(* IEC 61131-3 sources: SortJet_MasterSPS_Aufbau.fbsproj/Device.device.xml.v3^/Plc Logic.plclogic.xml.v3^/Application.application.xml.v3^/09_Station/Shuttle/[101,102] Shuttle/0_Konfig (part 2) *)

(* ---- Konfiguration_101.gvl ---- *)
(* METADATA
{
	"v3Meta": {
		"objectGuid": "a708fc7a-282c-4202-ac62-7eb4c755f260"
	}
}
*)
{attribute 'allow_unqualified_access'}
NAMESPACE Konfiguration_101
VAR_CONFIG
  // werden Variablen die gemappt werden hier ignoriert?
  // ------------------------------------------------- HARDWARE EINGAENGE -------------------------------------------------
  // Datenlichtschranke
  Globale_Bausteine.aShuttle[101].in_bDatenlichtschrankeShuttlebahnOK                                AT %MX1.1  : BOOL; // OPTION - Bauteil an der Shuttlebahn => Sender / Empfaenger
  Globale_Bausteine.aShuttle[101].in_bDatenlichtschrankeShuttleOK                                    AT %MX1.1  : BOOL; // OPTION - Bauteil auf dem Shuttle => Sender / Empfaenger

  // Sicherungen \ Motorschutzschalter \ etc.

  Globale_Bausteine.aShuttle[101].in_bSicherungen230V_OK                                             AT %MX1.1   : BOOL; // OPTION
  Globale_Bausteine.aShuttle[101].in_bLSQuerfahrtBremseOK                                            AT %IX101.0 : BOOL; // IO-L - Querfahrt Bremse Sicherung
  Globale_Bausteine.aShuttle[101].in_bNetzteil_24V_OK                                                AT %IX100.1 : BOOL; // IO-L - Netzteil 24V OK
  Globale_Bausteine.aShuttle[101].Kippen.in_bLeitungsschutzschalterBremseOK                          AT %MX1.1   : BOOL; // OPTION
  Globale_Bausteine.aShuttle[101].Kippen.in_bMotorschutzschalter_OK                                  AT %MX1.1   : BOOL; // OPTION

  // Druckluft
  Globale_Bausteine.aShuttle[101].in_bSicherungKompressor_OK                                         AT %MX1.1  : BOOL; // OPTION
  Globale_Bausteine.aShuttle[101].in_bDruckluft_OK                                                   AT %MX1.1  : BOOL; // OPTION

  //Geblaese Wand 1
  Globale_Bausteine.aShuttle[101].Geblaese[1].in_bMotorschutzschalter_OK                             AT %IX101.1  : BOOL; // IO-L - Geblaesegruppe Wand 1 Sicherung + Motorschutz
  Globale_Bausteine.aShuttle[101].Geblaese[1].out_bStarteGeblaese                                    AT %QX100.1  : BOOL; // IO-L - Geblaesegruppe Wand 1 einschalten

  // Wandverstellung Wand 1
  Globale_Bausteine.aShuttle[101].in_bWandverstellungsAntriebsSicherungOK                            AT %MX1.1   : BOOL; // OPTION
  Globale_Bausteine.aShuttle[101].in_bMotorstarterWandverstellungOK                                  AT %MX1.1   : BOOL; // OPTION
  Globale_Bausteine.aShuttle[101].in_bWandverstellungsBremsSicherungOK                               AT %MX1.1   : BOOL; // OPTION

  Globale_Bausteine.aShuttle[101].Wandverstellung[1].Pneumatik.in_bWandEinlaufseiteGeoeffnet         AT %MX1.0   : BOOL; // OPTION
  Globale_Bausteine.aShuttle[101].Wandverstellung[1].Pneumatik.in_bWandEinlaufseiteGeschlossen       AT %MX1.0   : BOOL; // OPTION
  Globale_Bausteine.aShuttle[101].Wandverstellung[1].Pneumatik.in_bWandAuslaufseiteGeoeffnet         AT %MX1.0   : BOOL; // OPTION
  Globale_Bausteine.aShuttle[101].Wandverstellung[1].Pneumatik.in_bWandAuslaufseiteGeschlossen       AT %MX1.0   : BOOL; // OPTION

  Globale_Bausteine.aShuttle[101].Wandverstellung[1].Pneumatik.out_bWandverstellungOeffnen           AT %MX1010.1 : BOOL; // OPTION
  Globale_Bausteine.aShuttle[101].Wandverstellung[1].Pneumatik.out_bWandverstellungSchliessen        AT %MX1010.2 : BOOL; // OPTION

  Globale_Bausteine.aShuttle[101].Wandverstellung[1].Pneumatik2.in_bStatusZylinder_Alle_Eingefahren  AT %MX1.0   : BOOL; // OPTION
  Globale_Bausteine.aShuttle[101].Wandverstellung[1].Pneumatik2.in_bStatusZylinder_1_Ausgefahren     AT %MX1.0   : BOOL; // OPTION
  Globale_Bausteine.aShuttle[101].Wandverstellung[1].Pneumatik2.in_bStatusZylinder_2_Ausgefahren     AT %MX1.0   : BOOL; // OPTION

  Globale_Bausteine.aShuttle[101].Wandverstellung[1].Pneumatik2.out_bZylinder_1_Einfahren            AT %MX1010.3 : BOOL; // OPTION
  Globale_Bausteine.aShuttle[101].Wandverstellung[1].Pneumatik2.out_bZylinder_2_Einfahren            AT %MX1010.4 : BOOL; // OPTION
  Globale_Bausteine.aShuttle[101].Wandverstellung[1].Pneumatik2.out_bZylinder_1_Ausfahren            AT %MX1010.5 : BOOL; // OPTION
  Globale_Bausteine.aShuttle[101].Wandverstellung[1].Pneumatik2.out_bZylinder_2_Ausfahren            AT %MX1010.6 : BOOL; // OPTION

  Globale_Bausteine.aShuttle[101].Wandverstellung[1].Rollenleiste.in_bStatusZylinder1Ausgefahren     AT %MX1.0   : BOOL; // OPTION
  Globale_Bausteine.aShuttle[101].Wandverstellung[1].Rollenleiste.in_bStatusZylinder1Eingefahren     AT %MX1.0   : BOOL; // OPTION
  Globale_Bausteine.aShuttle[101].Wandverstellung[1].Rollenleiste.in_bStatusZylinder2Ausgefahren     AT %MX1.0   : BOOL; // OPTION
  Globale_Bausteine.aShuttle[101].Wandverstellung[1].Rollenleiste.in_bStatusZylinder2Eingefahren     AT %MX1.0   : BOOL; // OPTION

  Globale_Bausteine.aShuttle[101].Wandverstellung[1].Rollenleiste.out_bZylinder1Einfahren            AT %MX1010.7 : BOOL; // OPTION
  Globale_Bausteine.aShuttle[101].Wandverstellung[1].Rollenleiste.out_bZylinder1Ausfahren            AT %MX1011.0 : BOOL; // OPTION
  Globale_Bausteine.aShuttle[101].Wandverstellung[1].Rollenleiste.out_bZylinder2Einfahren            AT %MX1011.1 : BOOL; // OPTION
  Globale_Bausteine.aShuttle[101].Wandverstellung[1].Rollenleiste.out_bZylinder2Ausfahren            AT %MX1011.2 : BOOL; // OPTION

  Globale_Bausteine.aShuttle[101].Wandverstellung[1].Rollenleiste_Schuetz.in_bVerstellungGeoeffnet   AT %MX1.0   : BOOL; // OPTION
  Globale_Bausteine.aShuttle[101].Wandverstellung[1].Rollenleiste_Schuetz.in_bVerstellungGeschlossen AT %MX1.0   : BOOL; // OPTION
  Globale_Bausteine.aShuttle[101].Wandverstellung[1].Rollenleiste_Schuetz.in_bMotorstarter_OK        AT %MX1.1   : BOOL; // OPTION
  Globale_Bausteine.aShuttle[101].Wandverstellung[1].Rollenleiste_Schuetz.in_bSicherungMotorOK       AT %MX1.1   : BOOL; // OPTION
  Globale_Bausteine.aShuttle[101].Wandverstellung[1].Rollenleiste_Schuetz.in_bBremseOK               AT %MX1.1   : BOOL; // OPTION

  Globale_Bausteine.aShuttle[101].Wandverstellung[1].Rollenleiste_Schuetz.out_bVerstellungSchliessen AT %MX1011.3 : BOOL; // OPTION
  Globale_Bausteine.aShuttle[101].Wandverstellung[1].Rollenleiste_Schuetz.out_bVerstellungOeffnen    AT %MX1011.4 : BOOL; // OPTION
  Globale_Bausteine.aShuttle[101].Wandverstellung[1].Rollenleiste_Schuetz.out_bBremseOeffnen         AT %MX1011.5 : BOOL; // OPTION
  Globale_Bausteine.aShuttle[101].Wandverstellung[1].Rollenleiste_Schuetz.out_bMotorstarterReset     AT %MX1011.6 : BOOL; // OPTION

  Globale_Bausteine.aShuttle[101].Wandverstellung[1].Gegenhalter_Schuetz.in_bVerstellungGeoeffnet    AT %MX1.0   : BOOL; // OPTION
  Globale_Bausteine.aShuttle[101].Wandverstellung[1].Gegenhalter_Schuetz.in_bVerstellungGeschlossen  AT %MX1.0   : BOOL; // OPTION
  Globale_Bausteine.aShuttle[101].Wandverstellung[1].Gegenhalter_Schuetz.in_bMotorstarter_OK         AT %MX1.1   : BOOL; // OPTION
  Globale_Bausteine.aShuttle[101].Wandverstellung[1].Gegenhalter_Schuetz.in_bSicherungMotorOK        AT %MX1.1   : BOOL; // OPTION
  Globale_Bausteine.aShuttle[101].Wandverstellung[1].Gegenhalter_Schuetz.in_bBremseOK                AT %MX1.1   : BOOL; // OPTION

  Globale_Bausteine.aShuttle[101].Wandverstellung[1].Gegenhalter_Schuetz.out_bVerstellungSchliessen  AT %MX1011.7 : BOOL; // OPTION
  Globale_Bausteine.aShuttle[101].Wandverstellung[1].Gegenhalter_Schuetz.out_bVerstellungOeffnen     AT %MX1012.0 : BOOL; // OPTION
  Globale_Bausteine.aShuttle[101].Wandverstellung[1].Gegenhalter_Schuetz.out_bBremseOeffnen          AT %MX1012.1 : BOOL; // OPTION
  Globale_Bausteine.aShuttle[101].Wandverstellung[1].Gegenhalter_Schuetz.out_bMotorstarterReset      AT %MX1012.2 : BOOL; // OPTION

  // Sensoren  Wand 2
  Globale_Bausteine.aShuttle[101].in_bSensorEinlaufVorabWand2                                        AT %MX1.0   : BOOL; // OPTION
  Globale_Bausteine.aShuttle[101].in_bSensorAuslaufVorabWand2                                        AT %MX1.0   : BOOL; // OPTION
  Globale_Bausteine.aShuttle[101].in_bSensorAuslaufStoppWand2                                        AT %MX1.0   : BOOL; // OPTION

  // Greifer Wand 1 [Ausbaustufe stStationsAufbau.bGreifer] (Kanaele laut Schaltplan eintragen, Glasrueckhalter laut Parameter_Greifer, ohne Bauteil Eingang auf %MX1.1)
  Globale_Bausteine.aShuttle[101].Greifer[1].in_bGreiferAusgefahren                                     AT %MX1.0   : BOOL; // OPTION
  Globale_Bausteine.aShuttle[101].Greifer[1].in_bGreiferEingefahren                                     AT %MX1.0   : BOOL; // OPTION
  Globale_Bausteine.aShuttle[101].Greifer[1].in_bGlasRueckhalterEinlaufEingefahren                      AT %MX1.1   : BOOL; // OPTION
  Globale_Bausteine.aShuttle[101].Greifer[1].in_bGlasRueckhalterAuslaufEingefahren                      AT %MX1.1   : BOOL; // OPTION

  Globale_Bausteine.aShuttle[101].Greifer[1].out_bGreiferAusfahren                                      AT %MX1012.3 : BOOL; // OPTION
  Globale_Bausteine.aShuttle[101].Greifer[1].out_bGreiferEinfahren                                      AT %MX1012.4 : BOOL; // OPTION
  Globale_Bausteine.aShuttle[101].Greifer[1].out_bGlasRueckhalterEinlaufAusfahren                       AT %MX1012.5 : BOOL; // OPTION
  Globale_Bausteine.aShuttle[101].Greifer[1].out_bGlasRueckhalterAuslaufAusfahren                       AT %MX1012.6 : BOOL; // OPTION

  // Greiferzange Einlaufseite Wand 1 [nur mit Parameter_Greifer.bZangeEinlaufVorhanden]
  Globale_Bausteine.aShuttle[101].Greifer[1].Zange[1].in_bStatusZylinder_Alle_Eingefahren               AT %MX1.0   : BOOL; // OPTION
  Globale_Bausteine.aShuttle[101].Greifer[1].Zange[1].in_bStatusZylinder_1_Ausgefahren                  AT %MX1.0   : BOOL; // OPTION
  Globale_Bausteine.aShuttle[101].Greifer[1].Zange[1].in_bStatusZylinder_2_Ausgefahren                  AT %MX1.0   : BOOL; // OPTION
  Globale_Bausteine.aShuttle[101].Greifer[1].Zange[1].in_bStatusZylinder_3_Ausgefahren                  AT %MX1.0   : BOOL; // OPTION

  Globale_Bausteine.aShuttle[101].Greifer[1].Zange[1].out_bZylinder_1_Einfahren                         AT %MX1012.7 : BOOL; // OPTION
  Globale_Bausteine.aShuttle[101].Greifer[1].Zange[1].out_bZylinder_2_Einfahren                         AT %MX1013.0 : BOOL; // OPTION
  Globale_Bausteine.aShuttle[101].Greifer[1].Zange[1].out_bZylinder_3_Einfahren                         AT %MX1013.1 : BOOL; // OPTION
  Globale_Bausteine.aShuttle[101].Greifer[1].Zange[1].out_bZylinder_1_Ausfahren                         AT %MX1013.2 : BOOL; // OPTION
  Globale_Bausteine.aShuttle[101].Greifer[1].Zange[1].out_bZylinder_2_Ausfahren                         AT %MX1013.3 : BOOL; // OPTION
  Globale_Bausteine.aShuttle[101].Greifer[1].Zange[1].out_bZylinder_3_Ausfahren                         AT %MX1013.4 : BOOL; // OPTION

  // Greiferzange Auslaufseite Wand 1 [nur mit Parameter_Greifer.bZangeAuslaufVorhanden]
  Globale_Bausteine.aShuttle[101].Greifer[1].Zange[2].in_bStatusZylinder_Alle_Eingefahren               AT %MX1.0   : BOOL; // OPTION
  Globale_Bausteine.aShuttle[101].Greifer[1].Zange[2].in_bStatusZylinder_1_Ausgefahren                  AT %MX1.0   : BOOL; // OPTION
  Globale_Bausteine.aShuttle[101].Greifer[1].Zange[2].in_bStatusZylinder_2_Ausgefahren                  AT %MX1.0   : BOOL; // OPTION
  Globale_Bausteine.aShuttle[101].Greifer[1].Zange[2].in_bStatusZylinder_3_Ausgefahren                  AT %MX1.0   : BOOL; // OPTION

  Globale_Bausteine.aShuttle[101].Greifer[1].Zange[2].out_bZylinder_1_Einfahren                         AT %MX1013.5 : BOOL; // OPTION
  Globale_Bausteine.aShuttle[101].Greifer[1].Zange[2].out_bZylinder_2_Einfahren                         AT %MX1013.6 : BOOL; // OPTION
  Globale_Bausteine.aShuttle[101].Greifer[1].Zange[2].out_bZylinder_3_Einfahren                         AT %MX1013.7 : BOOL; // OPTION
  Globale_Bausteine.aShuttle[101].Greifer[1].Zange[2].out_bZylinder_1_Ausfahren                         AT %MX1014.0 : BOOL; // OPTION
  Globale_Bausteine.aShuttle[101].Greifer[1].Zange[2].out_bZylinder_2_Ausfahren                         AT %MX1014.1 : BOOL; // OPTION
  Globale_Bausteine.aShuttle[101].Greifer[1].Zange[2].out_bZylinder_3_Ausfahren                         AT %MX1014.2 : BOOL; // OPTION

END_VAR

END_NAMESPACE

(* ---- Konfiguration_102.gvl ---- *)
(* METADATA
{
	"v3Meta": {
		"objectGuid": "12c6a77b-9420-47d5-ba1c-b94e93a145ed"
	}
}
*)
{attribute 'allow_unqualified_access'}
NAMESPACE Konfiguration_102
VAR_CONFIG
  // werden Variablen die gemappt werden hier ignoriert?
  // ------------------------------------------------- HARDWARE EINGAENGE -------------------------------------------------
  // Datenlichtschranke
  Globale_Bausteine.aShuttle[102].in_bDatenlichtschrankeShuttlebahnOK                                AT %MX1.1  : BOOL; // OPTION - Bauteil an der Shuttlebahn => Sender / Empfaenger
  Globale_Bausteine.aShuttle[102].in_bDatenlichtschrankeShuttleOK                                    AT %MX1.1  : BOOL; // OPTION - Bauteil auf dem Shuttle => Sender / Empfaenger

  // Sicherungen \ Motorschutzschalter \ etc.
  Globale_Bausteine.aShuttle[102].in_bSicherungen230V_OK                                             AT %MX1.1    : BOOL; // OPTION
  Globale_Bausteine.aShuttle[102].in_bLSQuerfahrtBremseOK                                            AT %IX111.0  : BOOL; // IO-L - Querfahrt Bremse Sicherung
  Globale_Bausteine.aShuttle[102].in_bNetzteil_24V_OK                                                AT %IX110.1  : BOOL; // IO-L - Netzteil 24V OK

  Globale_Bausteine.aShuttle[102].Kippen.in_bMotorschutzschalter_OK                                  AT %MX1.1   : BOOL; // OPTION
  Globale_Bausteine.aShuttle[102].Kippen.in_bLeitungsschutzschalterBremseOK                          AT %MX1.1   : BOOL; // OPTION

  // Druckluft
  Globale_Bausteine.aShuttle[102].in_bSicherungKompressor_OK                                         AT %MX1.1   : BOOL; // OPTION
  Globale_Bausteine.aShuttle[102].in_bDruckluft_OK                                                   AT %IX114.5 : BOOL; // IO-L - Druckluft OK

  //Geblaese Wand 1
  Globale_Bausteine.aShuttle[102].Geblaese[1].in_bMotorschutzschalter_OK                             AT %IX111.1  : BOOL; // IO-L - Geblaesegruppe Wand 1 Sicherung + Motorschutz
  Globale_Bausteine.aShuttle[102].Geblaese[1].out_bStarteGeblaese                                    AT %QX110.1  : BOOL; // IO-L - Geblaesegruppe Wand 1 einschalten

  // Wandverstellung Wand 1
  Globale_Bausteine.aShuttle[102].in_bWandverstellungsAntriebsSicherungOK                            AT %MX1.1   : BOOL; // OPTION
  Globale_Bausteine.aShuttle[102].in_bMotorstarterWandverstellungOK                                  AT %MX1.1   : BOOL; // OPTION
  Globale_Bausteine.aShuttle[102].in_bWandverstellungsBremsSicherungOK                               AT %MX1.1   : BOOL; // OPTION

  Globale_Bausteine.aShuttle[102].Wandverstellung[1].Pneumatik.in_bWandEinlaufseiteGeoeffnet         AT %MX1.0   : BOOL; // OPTION
  Globale_Bausteine.aShuttle[102].Wandverstellung[1].Pneumatik.in_bWandEinlaufseiteGeschlossen       AT %MX1.0   : BOOL; // OPTION
  Globale_Bausteine.aShuttle[102].Wandverstellung[1].Pneumatik.in_bWandAuslaufseiteGeoeffnet         AT %MX1.0   : BOOL; // OPTION
  Globale_Bausteine.aShuttle[102].Wandverstellung[1].Pneumatik.in_bWandAuslaufseiteGeschlossen       AT %MX1.0   : BOOL; // OPTION

  Globale_Bausteine.aShuttle[102].Wandverstellung[1].Pneumatik.out_bWandverstellungOeffnen           AT %MX1020.1 : BOOL; // OPTION
  Globale_Bausteine.aShuttle[102].Wandverstellung[1].Pneumatik.out_bWandverstellungSchliessen        AT %MX1020.2 : BOOL; // OPTION

  Globale_Bausteine.aShuttle[102].Wandverstellung[1].Pneumatik2.in_bStatusZylinder_Alle_Eingefahren  AT %MX1.0   : BOOL; // OPTION
  Globale_Bausteine.aShuttle[102].Wandverstellung[1].Pneumatik2.in_bStatusZylinder_1_Ausgefahren     AT %MX1.0   : BOOL; // OPTION
  Globale_Bausteine.aShuttle[102].Wandverstellung[1].Pneumatik2.in_bStatusZylinder_2_Ausgefahren     AT %MX1.0   : BOOL; // OPTION

  Globale_Bausteine.aShuttle[102].Wandverstellung[1].Pneumatik2.out_bZylinder_1_Einfahren            AT %MX1020.3 : BOOL; // OPTION
  Globale_Bausteine.aShuttle[102].Wandverstellung[1].Pneumatik2.out_bZylinder_2_Einfahren            AT %MX1020.4 : BOOL; // OPTION
  Globale_Bausteine.aShuttle[102].Wandverstellung[1].Pneumatik2.out_bZylinder_1_Ausfahren            AT %MX1020.5 : BOOL; // OPTION
  Globale_Bausteine.aShuttle[102].Wandverstellung[1].Pneumatik2.out_bZylinder_2_Ausfahren            AT %MX1020.6 : BOOL; // OPTION

  Globale_Bausteine.aShuttle[102].Wandverstellung[1].Rollenleiste.in_bStatusZylinder1Ausgefahren     AT %MX1.0   : BOOL; // OPTION
  Globale_Bausteine.aShuttle[102].Wandverstellung[1].Rollenleiste.in_bStatusZylinder1Eingefahren     AT %MX1.0   : BOOL; // OPTION
  Globale_Bausteine.aShuttle[102].Wandverstellung[1].Rollenleiste.in_bStatusZylinder2Ausgefahren     AT %MX1.0   : BOOL; // OPTION
  Globale_Bausteine.aShuttle[102].Wandverstellung[1].Rollenleiste.in_bStatusZylinder2Eingefahren     AT %MX1.0   : BOOL; // OPTION

  Globale_Bausteine.aShuttle[102].Wandverstellung[1].Rollenleiste.out_bZylinder1Einfahren            AT %MX1020.7 : BOOL; // OPTION
  Globale_Bausteine.aShuttle[102].Wandverstellung[1].Rollenleiste.out_bZylinder1Ausfahren            AT %MX1021.0 : BOOL; // OPTION
  Globale_Bausteine.aShuttle[102].Wandverstellung[1].Rollenleiste.out_bZylinder2Einfahren            AT %MX1021.1 : BOOL; // OPTION
  Globale_Bausteine.aShuttle[102].Wandverstellung[1].Rollenleiste.out_bZylinder2Ausfahren            AT %MX1021.2 : BOOL; // OPTION

  Globale_Bausteine.aShuttle[102].Wandverstellung[1].Rollenleiste_Schuetz.in_bVerstellungGeoeffnet   AT %MX1.0   : BOOL; // OPTION
  Globale_Bausteine.aShuttle[102].Wandverstellung[1].Rollenleiste_Schuetz.in_bVerstellungGeschlossen AT %MX1.0   : BOOL; // OPTION
  Globale_Bausteine.aShuttle[102].Wandverstellung[1].Rollenleiste_Schuetz.in_bMotorstarter_OK        AT %MX1.1   : BOOL; // OPTION
  Globale_Bausteine.aShuttle[102].Wandverstellung[1].Rollenleiste_Schuetz.in_bSicherungMotorOK       AT %MX1.1   : BOOL; // OPTION
  Globale_Bausteine.aShuttle[102].Wandverstellung[1].Rollenleiste_Schuetz.in_bBremseOK               AT %MX1.1   : BOOL; // OPTION

  Globale_Bausteine.aShuttle[102].Wandverstellung[1].Rollenleiste_Schuetz.out_bVerstellungSchliessen AT %MX1021.3 : BOOL; // OPTION
  Globale_Bausteine.aShuttle[102].Wandverstellung[1].Rollenleiste_Schuetz.out_bVerstellungOeffnen    AT %MX1021.4 : BOOL; // OPTION
  Globale_Bausteine.aShuttle[102].Wandverstellung[1].Rollenleiste_Schuetz.out_bBremseOeffnen         AT %MX1021.5 : BOOL; // OPTION
  Globale_Bausteine.aShuttle[102].Wandverstellung[1].Rollenleiste_Schuetz.out_bMotorstarterReset     AT %MX1021.6 : BOOL; // OPTION

  Globale_Bausteine.aShuttle[102].Wandverstellung[1].Gegenhalter_Schuetz.in_bVerstellungGeoeffnet    AT %MX1.0   : BOOL; // OPTION
  Globale_Bausteine.aShuttle[102].Wandverstellung[1].Gegenhalter_Schuetz.in_bVerstellungGeschlossen  AT %MX1.0   : BOOL; // OPTION
  Globale_Bausteine.aShuttle[102].Wandverstellung[1].Gegenhalter_Schuetz.in_bMotorstarter_OK         AT %MX1.1   : BOOL; // OPTION
  Globale_Bausteine.aShuttle[102].Wandverstellung[1].Gegenhalter_Schuetz.in_bSicherungMotorOK        AT %MX1.1   : BOOL; // OPTION
  Globale_Bausteine.aShuttle[102].Wandverstellung[1].Gegenhalter_Schuetz.in_bBremseOK                AT %MX1.1   : BOOL; // OPTION

  Globale_Bausteine.aShuttle[102].Wandverstellung[1].Gegenhalter_Schuetz.out_bVerstellungSchliessen  AT %MX1021.7 : BOOL; // OPTION
  Globale_Bausteine.aShuttle[102].Wandverstellung[1].Gegenhalter_Schuetz.out_bVerstellungOeffnen     AT %MX1022.0 : BOOL; // OPTION
  Globale_Bausteine.aShuttle[102].Wandverstellung[1].Gegenhalter_Schuetz.out_bBremseOeffnen          AT %MX1022.1 : BOOL; // OPTION
  Globale_Bausteine.aShuttle[102].Wandverstellung[1].Gegenhalter_Schuetz.out_bMotorstarterReset      AT %MX1022.2 : BOOL; // OPTION

  // Sensoren  Wand 2
  Globale_Bausteine.aShuttle[102].in_bSensorEinlaufVorabWand2                                        AT %MX1.0   : BOOL; // OPTION
  Globale_Bausteine.aShuttle[102].in_bSensorAuslaufVorabWand2                                        AT %MX1.0   : BOOL; // OPTION
  Globale_Bausteine.aShuttle[102].in_bSensorAuslaufStoppWand2                                        AT %MX1.0   : BOOL; // OPTION

  //Geblaese Wand 2
  Globale_Bausteine.aShuttle[102].Geblaese[2].in_bMotorschutzschalter_OK                             AT %MX1.1    : BOOL; // OPTION
  Globale_Bausteine.aShuttle[102].Geblaese[2].out_bStarteGeblaese                                    AT %MX1022.3 : BOOL; // OPTION

  // Wandverstellung Wand 2
  Globale_Bausteine.aShuttle[102].Wandverstellung[2].Pneumatik.in_bWandEinlaufseiteGeoeffnet         AT %MX1.0   : BOOL; // OPTION
  Globale_Bausteine.aShuttle[102].Wandverstellung[2].Pneumatik.in_bWandEinlaufseiteGeschlossen       AT %MX1.0   : BOOL; // OPTION
  Globale_Bausteine.aShuttle[102].Wandverstellung[2].Pneumatik.in_bWandAuslaufseiteGeoeffnet         AT %MX1.0   : BOOL; // OPTION
  Globale_Bausteine.aShuttle[102].Wandverstellung[2].Pneumatik.in_bWandAuslaufseiteGeschlossen       AT %MX1.0   : BOOL; // OPTION

  Globale_Bausteine.aShuttle[102].Wandverstellung[2].Pneumatik.out_bWandverstellungOeffnen           AT %MX1022.4 : BOOL; // OPTION
  Globale_Bausteine.aShuttle[102].Wandverstellung[2].Pneumatik.out_bWandverstellungSchliessen        AT %MX1022.5 : BOOL; // OPTION

  Globale_Bausteine.aShuttle[102].Wandverstellung[2].Pneumatik2.in_bStatusZylinder_Alle_Eingefahren  AT %MX1.0   : BOOL; // OPTION
  Globale_Bausteine.aShuttle[102].Wandverstellung[2].Pneumatik2.in_bStatusZylinder_1_Ausgefahren     AT %MX1.0   : BOOL; // OPTION
  Globale_Bausteine.aShuttle[102].Wandverstellung[2].Pneumatik2.in_bStatusZylinder_2_Ausgefahren     AT %MX1.0   : BOOL; // OPTION

  Globale_Bausteine.aShuttle[102].Wandverstellung[2].Pneumatik2.out_bZylinder_1_Einfahren            AT %MX1022.6 : BOOL; // OPTION
  Globale_Bausteine.aShuttle[102].Wandverstellung[2].Pneumatik2.out_bZylinder_2_Einfahren            AT %MX1022.7 : BOOL; // OPTION
  Globale_Bausteine.aShuttle[102].Wandverstellung[2].Pneumatik2.out_bZylinder_1_Ausfahren            AT %MX1023.0 : BOOL; // OPTION
  Globale_Bausteine.aShuttle[102].Wandverstellung[2].Pneumatik2.out_bZylinder_2_Ausfahren            AT %MX1023.1 : BOOL; // OPTION

  Globale_Bausteine.aShuttle[102].Wandverstellung[2].Rollenleiste.in_bStatusZylinder1Ausgefahren     AT %MX1.0   : BOOL; // OPTION
  Globale_Bausteine.aShuttle[102].Wandverstellung[2].Rollenleiste.in_bStatusZylinder1Eingefahren     AT %MX1.0   : BOOL; // OPTION
  Globale_Bausteine.aShuttle[102].Wandverstellung[2].Rollenleiste.in_bStatusZylinder2Ausgefahren     AT %MX1.0   : BOOL; // OPTION
  Globale_Bausteine.aShuttle[102].Wandverstellung[2].Rollenleiste.in_bStatusZylinder2Eingefahren     AT %MX1.0   : BOOL; // OPTION

  Globale_Bausteine.aShuttle[102].Wandverstellung[2].Rollenleiste.out_bZylinder1Einfahren            AT %MX1023.2 : BOOL; // OPTION
  Globale_Bausteine.aShuttle[102].Wandverstellung[2].Rollenleiste.out_bZylinder1Ausfahren            AT %MX1023.3 : BOOL; // OPTION
  Globale_Bausteine.aShuttle[102].Wandverstellung[2].Rollenleiste.out_bZylinder2Einfahren            AT %MX1023.4 : BOOL; // OPTION
  Globale_Bausteine.aShuttle[102].Wandverstellung[2].Rollenleiste.out_bZylinder2Ausfahren            AT %MX1023.5 : BOOL; // OPTION

  Globale_Bausteine.aShuttle[102].Wandverstellung[2].Rollenleiste_Schuetz.in_bVerstellungGeoeffnet   AT %MX1.0   : BOOL; // OPTION
  Globale_Bausteine.aShuttle[102].Wandverstellung[2].Rollenleiste_Schuetz.in_bVerstellungGeschlossen AT %MX1.0   : BOOL; // OPTION
  Globale_Bausteine.aShuttle[102].Wandverstellung[2].Rollenleiste_Schuetz.in_bMotorstarter_OK        AT %MX1.1   : BOOL; // OPTION
  Globale_Bausteine.aShuttle[102].Wandverstellung[2].Rollenleiste_Schuetz.in_bSicherungMotorOK       AT %MX1.1   : BOOL; // OPTION
  Globale_Bausteine.aShuttle[102].Wandverstellung[2].Rollenleiste_Schuetz.in_bBremseOK               AT %MX1.1   : BOOL; // OPTION

  Globale_Bausteine.aShuttle[102].Wandverstellung[2].Rollenleiste_Schuetz.out_bVerstellungSchliessen AT %MX1023.6 : BOOL; // OPTION
  Globale_Bausteine.aShuttle[102].Wandverstellung[2].Rollenleiste_Schuetz.out_bVerstellungOeffnen    AT %MX1023.7 : BOOL; // OPTION
  Globale_Bausteine.aShuttle[102].Wandverstellung[2].Rollenleiste_Schuetz.out_bBremseOeffnen         AT %MX1024.0 : BOOL; // OPTION
  Globale_Bausteine.aShuttle[102].Wandverstellung[2].Rollenleiste_Schuetz.out_bMotorstarterReset     AT %MX1024.1 : BOOL; // OPTION

  Globale_Bausteine.aShuttle[102].Wandverstellung[2].Gegenhalter_Schuetz.in_bVerstellungGeoeffnet    AT %MX1.0   : BOOL; // OPTION
  Globale_Bausteine.aShuttle[102].Wandverstellung[2].Gegenhalter_Schuetz.in_bVerstellungGeschlossen  AT %MX1.0   : BOOL; // OPTION
  Globale_Bausteine.aShuttle[102].Wandverstellung[2].Gegenhalter_Schuetz.in_bMotorstarter_OK         AT %MX1.1   : BOOL; // OPTION
  Globale_Bausteine.aShuttle[102].Wandverstellung[2].Gegenhalter_Schuetz.in_bSicherungMotorOK        AT %MX1.1   : BOOL; // OPTION
  Globale_Bausteine.aShuttle[102].Wandverstellung[2].Gegenhalter_Schuetz.in_bBremseOK                AT %MX1.1   : BOOL; // OPTION

  Globale_Bausteine.aShuttle[102].Wandverstellung[2].Gegenhalter_Schuetz.out_bVerstellungSchliessen  AT %MX1024.2 : BOOL; // OPTION
  Globale_Bausteine.aShuttle[102].Wandverstellung[2].Gegenhalter_Schuetz.out_bVerstellungOeffnen     AT %MX1024.3 : BOOL; // OPTION
  Globale_Bausteine.aShuttle[102].Wandverstellung[2].Gegenhalter_Schuetz.out_bBremseOeffnen          AT %MX1024.4 : BOOL; // OPTION
  Globale_Bausteine.aShuttle[102].Wandverstellung[2].Gegenhalter_Schuetz.out_bMotorstarterReset      AT %MX1024.5 : BOOL; // OPTION

  // Greifer Wand 1 [Ausbaustufe stStationsAufbau.bGreifer] (Kanaele laut Schaltplan eintragen, Glasrueckhalter laut Parameter_Greifer, ohne Bauteil Eingang auf %MX1.1)
  Globale_Bausteine.aShuttle[102].Greifer[1].in_bGreiferAusgefahren                                     AT %IX113.0  : BOOL; // IO-L - Greifer 1 ausgefahren zum Glas
  Globale_Bausteine.aShuttle[102].Greifer[1].in_bGreiferEingefahren                                     AT %IX113.1  : BOOL; // IO-L - Greifer 1 eingefahren
  Globale_Bausteine.aShuttle[102].Greifer[1].in_bGlasRueckhalterEinlaufEingefahren                      AT %MX1.1    : BOOL; // OPTION - Einlaufseite ohne Glasrueckhalter
  Globale_Bausteine.aShuttle[102].Greifer[1].in_bGlasRueckhalterAuslaufEingefahren                      AT %IX113.4  : BOOL; // IO-L - Greifer 1 Haltebuegel eingefahren

  Globale_Bausteine.aShuttle[102].Greifer[1].out_bGreiferAusfahren                                      AT %QX110.7   : BOOL; // IO-L - Greifer 1 ausfahren zum Glas
  Globale_Bausteine.aShuttle[102].Greifer[1].out_bGreiferEinfahren                                      AT %QX111.0   : BOOL; // IO-L - Greifer 1 einfahren
  Globale_Bausteine.aShuttle[102].Greifer[1].out_bGlasRueckhalterEinlaufAusfahren                       AT %MX1025.0  : BOOL; // OPTION
  Globale_Bausteine.aShuttle[102].Greifer[1].out_bGlasRueckhalterAuslaufAusfahren                       AT %QX111.3   : BOOL; // IO-L - Greifer 1 Haltebuegel ausfahren

  // Greiferzange Einlaufseite Wand 1 [nur mit Parameter_Greifer.bZangeEinlaufVorhanden]
  Globale_Bausteine.aShuttle[102].Greifer[1].Zange[1].in_bStatusZylinder_Alle_Eingefahren               AT %MX1.0   : BOOL; // OPTION
  Globale_Bausteine.aShuttle[102].Greifer[1].Zange[1].in_bStatusZylinder_1_Ausgefahren                  AT %MX1.0   : BOOL; // OPTION
  Globale_Bausteine.aShuttle[102].Greifer[1].Zange[1].in_bStatusZylinder_2_Ausgefahren                  AT %MX1.0   : BOOL; // OPTION
  Globale_Bausteine.aShuttle[102].Greifer[1].Zange[1].in_bStatusZylinder_3_Ausgefahren                  AT %MX1.0   : BOOL; // OPTION

  Globale_Bausteine.aShuttle[102].Greifer[1].Zange[1].out_bZylinder_1_Einfahren                         AT %MX1025.2 : BOOL; // OPTION
  Globale_Bausteine.aShuttle[102].Greifer[1].Zange[1].out_bZylinder_2_Einfahren                         AT %MX1025.3 : BOOL; // OPTION
  Globale_Bausteine.aShuttle[102].Greifer[1].Zange[1].out_bZylinder_3_Einfahren                         AT %MX1025.4 : BOOL; // OPTION
  Globale_Bausteine.aShuttle[102].Greifer[1].Zange[1].out_bZylinder_1_Ausfahren                         AT %MX1025.5 : BOOL; // OPTION
  Globale_Bausteine.aShuttle[102].Greifer[1].Zange[1].out_bZylinder_2_Ausfahren                         AT %MX1025.6 : BOOL; // OPTION
  Globale_Bausteine.aShuttle[102].Greifer[1].Zange[1].out_bZylinder_3_Ausfahren                         AT %MX1025.7 : BOOL; // OPTION

  // Greiferzange Auslaufseite Wand 1 [nur mit Parameter_Greifer.bZangeAuslaufVorhanden]
  Globale_Bausteine.aShuttle[102].Greifer[1].Zange[2].in_bStatusZylinder_Alle_Eingefahren               AT %IX113.2 : BOOL; // IO-L - Greifer 1 Hub 1 geschlossen (nicht ausgewertet, bZangeAbfragenVorhanden = FALSE)
  Globale_Bausteine.aShuttle[102].Greifer[1].Zange[2].in_bStatusZylinder_1_Ausgefahren                 AT %IX113.3 : BOOL; // IO-L - Greifer 1 Hub 1 geoeffnet
  Globale_Bausteine.aShuttle[102].Greifer[1].Zange[2].in_bStatusZylinder_2_Ausgefahren                  AT %MX1.0   : BOOL; // OPTION
  Globale_Bausteine.aShuttle[102].Greifer[1].Zange[2].in_bStatusZylinder_3_Ausgefahren                  AT %MX1.0   : BOOL; // OPTION

  Globale_Bausteine.aShuttle[102].Greifer[1].Zange[2].out_bZylinder_1_Einfahren                         AT %QX111.2  : BOOL; // IO-L - Greifer 1 Hub 1 schliessen
  Globale_Bausteine.aShuttle[102].Greifer[1].Zange[2].out_bZylinder_2_Einfahren                         AT %MX1026.1 : BOOL; // OPTION
  Globale_Bausteine.aShuttle[102].Greifer[1].Zange[2].out_bZylinder_3_Einfahren                         AT %MX1026.2 : BOOL; // OPTION
  Globale_Bausteine.aShuttle[102].Greifer[1].Zange[2].out_bZylinder_1_Ausfahren                         AT %QX111.1  : BOOL; // IO-L - Greifer 1 Hub 1 oeffnen
  Globale_Bausteine.aShuttle[102].Greifer[1].Zange[2].out_bZylinder_2_Ausfahren                         AT %MX1026.4 : BOOL; // OPTION
  Globale_Bausteine.aShuttle[102].Greifer[1].Zange[2].out_bZylinder_3_Ausfahren                         AT %MX1026.5 : BOOL; // OPTION

END_VAR

END_NAMESPACE

(* ---- Konfiguration_Optionales.gvl ---- *)
(* METADATA
{
	"v3Meta": {
		"objectGuid": "a15d5673-fc2e-4b3d-8d8d-59c1778f3865"
	}
}
*)
{attribute 'allow_unqualified_access'}
NAMESPACE Konfiguration_Optionales
VAR_CONFIG

  // Sensoren  Wand 2
  Globale_Bausteine.aShuttle[101].in_bSensorEinlaufVorabWand2                                        AT %MX1.0   : BOOL; // OPTION
  Globale_Bausteine.aShuttle[101].in_bSensorAuslaufVorabWand2                                        AT %MX1.0   : BOOL; // OPTION
  Globale_Bausteine.aShuttle[101].in_bSensorAuslaufStoppWand2                                        AT %MX1.0   : BOOL; // OPTION

  //Geblaese Wand 2
  Globale_Bausteine.aShuttle[101].Geblaese[2].in_bMotorschutzschalter_OK                             AT %MX1.1    : BOOL; // OPTION
  Globale_Bausteine.aShuttle[101].Geblaese[2].out_bStarteGeblaese                                    AT %MX920.0  : BOOL; // OPTION

  //Geblaese Wand 3
  Globale_Bausteine.aShuttle[101].Geblaese[3].in_bMotorschutzschalter_OK                             AT %MX1.1    : BOOL; // OPTION
  Globale_Bausteine.aShuttle[101].Geblaese[3].out_bStarteGeblaese                                    AT %MX920.1  : BOOL; // OPTION

END_VAR
END_NAMESPACE
